Fanuc KAREL source: KA00085.KL

PROGRAM KA00085
%NOLOCKGROUP
VAR
  SRC: JOINTPOS
  DST: INTEGER
BEGIN
  DST = SRC
END KA00085
